Staubli VAL3: HMI_pointEdit.dtx

mdesc mNomSpeed
bool bBack
string sTrajItem
string sUsingLib
string sUsingFrame
string sUsingTool
public bool bBool[30]
string sPageIndex
string sPageNum
public string sList = "0"
string sSelPoint
num nPageIndex
num nPageNum
bool bRefresh
bool bConfirm
bool bBackSignal
string sSignalType
string sSignalIndex
num nSignalValue
num nSignalType
string sLastType
string sIOList
bool bConfirmDelay
bool bBackDelay
num nSetDelay
public string sIFtype[3]
string sIFIndex[3]
public num nIOindex[3]
public num nIFvalue[3]
bool bConfirmIF
bool bBackIF
string sANDOR[2]
public num nANDOR[2]
num nIFtype[3]
num nParaSpeed
num nParaAccel
num nParaBlend
num nParaPercent
string sParaType
bool bParaJoint
bool bParaOFF
num nMoveType
bool bParaConfirm
bool bParaBack
bool bPAllModify
bool bLast
bool bToSave
frame fUsingFrame = {fatherId=world[0]}
tool tUsingTool = {fatherId=flange[0]}
public num nTRSF[12]
public string sTRSF[12]
string sBlendType
string sLastItem
string sLastMtype
num _nFrameID
num _nToolID
num _nPointIndex
string sComment
num nPointIndex
bool bSafePoint
string sActionList
bool bAConfirm
bool bACancel
string sSelAction
bool bConfirmSwitch
bool bBackSwitch
bool bMark
public string sCommentIO1
bool bToSave1
string sLastTrajItem
string sSelMovCPoint
bool bRecord
bool bMoveTo
bool bConfirmMovC
bool bCancelMovC
bool bShow2Point
string sParaPointType[2]
